(* IEC 61131-3 sources: plc-ci-toolkit/ci/tests/samples/sa_probe_src/src/POUs/PRG_SaTask2, 1 file *)

(* ---- PRG_SaTask2.decl.st ---- *)
// Назначение: зонд статанализа — вторая задача
PROGRAM PRG_SaTask2
VAR
END_VAR
